FUNCTION_BLOCK FINAL CM_ControlModule EXTENDS PML_Module IMPLEMENTS I_CmControlModule
VAR_IN_OUT
    DevList : ST_ControlModuleDevList;
END_VAR
VAR
	// Tags trailing properties


	// PB Instance Declaration


	// Sequence Instance Declaration
	seqModuleSequence	: SEQ_ModuleSequence := (Description := 'Module Sequence', _enableHmiStart := TRUE, _enableSfcTipCtrl := FALSE);

	// Module/Device Instance Declaration

	// Other local variables
	cmd	: E_CmControlModuleCmd;

END_VAR

// Call Pushbutton FBs (or Update command)


// Evaluate commands to drive states, run methods of devices (ax.MoveAbs), run seq etc.
StateTransitionLogic();

// Call Sequence FBs
// Call Sequence FBs
seqModuleSequence(DevList := THIS^.DevList);

// Call Module/Device FBs
SUPER^(); // Basically a module. Call other modules below this.


// Reset cmd at end of FB Scan
cmd := E_CmControlModuleCmd.NoCmd;

METHOD PRIVATE InitAlarms : BOOL
END_METHOD

METHOD PRIVATE RaiseAlarm : BOOL
VAR_INPUT
	AlarmId : UDINT;
END_VAR
CASE AlarmId OF
0:
	;
END_CASE
END_METHOD

METHOD PROTECTED RunPmlExecute
// Add custom implementation
CASE CurrentPmlMode OF
	E_PmlMode.Production:
		//

	E_PmlMode.SemiAuto:
		//

	E_PmlMode.Manual:
		//

END_CASE
END_METHOD

METHOD PROTECTED SetDependency
// Attach Sequences
Attach(seqModuleSequence);

// Attach Modules/Devices

// The warning can be disabled here as the user is aware of the risk that the reference may not be valid by checking its validity
{warning disable C0371}

// Checking the VAR_IN_OUT reference, leave the current method in case of invalid reference
IF NOT __ISVALIDREF(DevList) THEN
     RETURN;
END_IF

// Access to VAR_IN_OUT reference (only if the reference was confirmed as valid before)
AttachDevList(ListPointer := ADR(DevList), ListSize := SIZEOF(DevList));

// The warning may be restored at the end of the access area
{warning restore C0371}
SUPER^.SetDependency(); // Call at the end, after all of the attach
END_METHOD

METHOD PRIVATE StateTransitionLogic
END_METHOD

END_FUNCTION_BLOCK

(* stored: Version 1.1.0.1, ProductVersion 3.1.4024.12
   POU CM_ControlModule: Id {6bd9f387-eeb9-4515-9779-aa7709b1122b}, SpecialFunc None
   Folder Interface Methods: Id {07c18477-deb2-4f8f-8bb0-9f2f98c77fae}
   Folder Interface Properties: Id {b53d5b70-581e-47aa-8ccc-d349c865956c}
   Folder PBs: Id {2415b04f-52f8-46fe-aae2-14920befeb5b}
   Folder Override Methods: Id {f166f506-d564-48b0-bc0b-d85579121499}
   Folder Alarm Methods: Id {67d5975e-da59-41cd-9e2b-c649c072069f}
   Folder PML State Methods: Id {207ce5fe-9b50-4b4f-8d5e-18c54ee32d60}
   Folder Override Properties: Id {f4d0ca19-06ae-4acb-9cf0-8e582dd7d3a4}
   Folder PBs: Id {41b8106d-78c5-45f8-a060-b726c2df9a8b}
   Folder Private Methods: Id {df29cb4e-1f08-4ac4-b495-c7ec4478b825}
   Method InitAlarms: Id {536445a3-f197-4bc3-a73f-5691a2fa7e9e}
   Method RaiseAlarm: Id {6eefa232-6459-4c40-a7f0-20ed389d05a0}
   Method RunPmlExecute: Id {d0d30f7a-bdd3-450c-8e7d-1d3fbeb1edbb}
   Method SetDependency: Id {35445cbb-64bd-4192-bb62-69b56d940994}
   Method StateTransitionLogic: Id {34a273d8-4104-4c06-9c03-b4f26a86d847} *)
